(* PLC project PumpStation, Example Water Co. CODESYS CODESYS V3.5 SP19 *)
(* stored: creationDateTime 2026-11-16T09:00:00, modificationDateTime 2026-11-16T09:00:00 *)

TYPE E_PumpState : (Idle := 0, Running := 1, Faulted := 2);
END_TYPE

TYPE ST_Pump : STRUCT
  State : E_PumpState;
  Speed : REAL;  (* Speed in percent *)
  Hours : UDINT;
END_STRUCT;
END_TYPE

(* Level-controlled pump with hysteresis *)
FUNCTION_BLOCK FB_Pump
  VAR_INPUT
    xEnable : BOOL;
    rLevel : REAL;  (* Tank level in m *)
  END_VAR
  VAR_OUTPUT
    xRun : BOOL;
  END_VAR
  VAR CONSTANT
    START_LEVEL : REAL := 2.5;
    STOP_LEVEL : REAL := 0.8;
  END_VAR

            IF NOT xEnable THEN
    xRun := FALSE;
ELSIF rLevel > START_LEVEL THEN
    xRun := TRUE;
ELSIF rLevel < STOP_LEVEL THEN
    xRun := FALSE;
END_IF
          
END_FUNCTION_BLOCK

PROGRAM PLC_PRG
  VAR
    fbPump1 : FB_Pump;
    aLevels : ARRAY[1..4] OF REAL;
  END_VAR

            fbPump1(xEnable := GVL.xAuto, rLevel := aLevels[1]);
GVL.xPump1Run := fbPump1.xRun;
          
END_PROGRAM

PROGRAM Alarms
  VAR
    xHighLevel : BOOL;
  END_VAR

(* LD diagram, written out as Structured Text *)
xHighLevel := GVL.xLevelHighSwitch;
END_PROGRAM

CONFIGURATION Device
  RESOURCE Application ON PLC
    VAR_GLOBAL  (* GVL *)
      xAuto : BOOL := TRUE;
      xPump1Run AT %QX0.0 : BOOL;
      xLevelHighSwitch AT %IX0.3 : BOOL;
    END_VAR
    TASK MainTask(INTERVAL := T#20ms, PRIORITY := 1);
    PROGRAM PLC_PRG WITH MainTask : PLC_PRG;
    PROGRAM Alarms WITH MainTask : Alarms;
  END_RESOURCE
END_CONFIGURATION
